FUNCTION_BLOCK Controle_Necessidade_HMI (* Service Interface Function Block Type *)
  (* Standard: 61499-2 *)
  (* Version 1.0, 21/10/2026, Hidryco, Hidryco, IHM do Controle_Necessidade *)
  PACKAGE Hidryco.HidrycoLib;
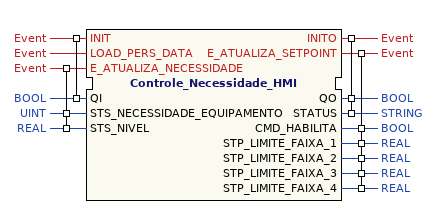
  EVENT_INPUT
    INIT WITH QI;
    LOAD_PERS_DATA; (* Reenvia os parametros persistentes *)
    E_ATUALIZA_NECESSIDADE WITH STS_NECESSIDADE_EQUIPAMENTO, STS_NIVEL; (* Status do processo *)
  END_EVENT
  EVENT_OUTPUT
    INITO WITH QO, STATUS;
    E_ATUALIZA_SETPOINT WITH STP_LIMITE_FAIXA_1, STP_LIMITE_FAIXA_2, STP_LIMITE_FAIXA_3, STP_LIMITE_FAIXA_4, CMD_HABILITA; (* Ajustes (IHM/OPC UA e LOAD_PERS_DATA) *)
  END_EVENT
  VAR_INPUT
    QI : BOOL;
    STS_NECESSIDADE_EQUIPAMENTO : UINT; (* Equipamentos pedidos pelas faixas *)
    STS_NIVEL : REAL; (* Nivel comparado com as faixas (% da altura) *)
  END_VAR
  VAR_OUTPUT
    QO : BOOL; (* Event Output Qualifier *)
    STATUS : STRING; (* Service Status *)
    CMD_HABILITA : BOOL; (* Habilitado *)
    STP_LIMITE_FAIXA_1 : REAL; (* Limite da faixa 1 *)
    STP_LIMITE_FAIXA_2 : REAL; (* Limite da faixa 2 *)
    STP_LIMITE_FAIXA_3 : REAL; (* Limite da faixa 3 *)
    STP_LIMITE_FAIXA_4 : REAL; (* Limite da faixa 4 *)
  END_VAR
  SERVICE /
    SEQUENCE 
    END_SEQUENCE
  END_SERVICE
END_FUNCTION_BLOCK
